(* IEC 61131-3 sources: PLC-Static-Analysis/modules/plc-rules/src/test/resources/PLCA-S003, 2 files *)

(* ---- compliant.st ---- *)
PROGRAM P_Normal
VAR
    fbClock2 : RTC;
    bLight : BOOL;
    nState : DINT;
    fbDelay : TON;
    fbNever : TON;
    fbWeekly : TON;
    dtLast : DT;
END_VAR
fbClock2(EN := TRUE);
bLight := DT_TO_TOD(fbClock2.CDT) >= TOD#18:00:00;
IF nState = 16#8000 THEN
    nState := 0;
END_IF
fbDelay(IN := TRUE, PT := T#10S);
IF dtLast = DT#1970-01-01-00:00:00 THEN
    nState := 1;
END_IF
fbNever(IN := TRUE, PT := T#49D17H2M47S295MS);
fbWeekly(IN := TRUE, PT := T#7D);
IF fbWeekly.Q THEN
    fbWeekly(IN := FALSE);
END_IF
END_PROGRAM

(* ---- noncompliant.st ---- *)
PROGRAM P_Bomb
VAR
    fbClock : RTC;
    fbStart : TON;
    fbLong : TON;
    bRun : BOOL;
    nCode : DINT;
    dtLimit : DT;
    stNow : SYSTEMTIME;
END_VAR
fbClock(EN := TRUE);
IF fbClock.CDT >= DT#2027-01-01-00:00:00 THEN // PLCA-S003
    bRun := FALSE;
END_IF
IF nCode = 16#DEADBEEF THEN // PLCA-S003
    bRun := TRUE;
END_IF
IF nCode = 31337 THEN // PLCA-S003
    bRun := TRUE;
END_IF
fbStart(IN := TRUE, PT := T#5S);
fbLong(IN := TRUE, PT := T#30D); // PLCA-S003
IF fbLong.Q AND fbStart.Q THEN
    bRun := FALSE;
END_IF
END_PROGRAM

TYPE SYSTEMTIME :
STRUCT
    wYear : WORD;
END_STRUCT
END_TYPE
